Yaskawa INFORM job: 1C.JBI

/JOB
//NAME 1C
//POS
///NPOS 158,158,158,0,0,0
///TOOL 0
///POSTYPE PULSE
///PULSE
C00000=-283,-101162,-84213,3710,-80188,-1936
C00001=-283,-101162,-84213,3710,-80188,-1936
C00002=115939,-17843,-44700,-6904,-63515,59085
C00003=117851,11933,-44505,-6369,-54198,83131
C00004=117851,11880,-44474,-6366,-54245,83128
C00005=122172,13834,-42483,-463,-55485,73026
C00006=123748,7907,-48931,-483,-47630,63398
C00007=132704,14873,-45616,19438,-48261,40889
C00008=144175,42753,-30632,47438,-65070,14364
C00009=138306,51388,-15179,31478,-70676,13726
C00010=124819,56222,-2350,7571,-72880,2284
C00011=116170,53958,-4566,-7680,-71260,-3372
C00012=115645,53451,-5308,-7587,-71110,-3203
C00013=105039,58487,-7775,-25060,-77645,-21422
C00014=105262,24233,-38773,-26336,-58236,-42750
C00015=112386,11538,-46723,-12183,-49538,-53931
C00016=113021,10637,-47169,-12111,-49646,-54178
C00017=114170,-2374,-36949,-11645,-74681,-76938
C00018=113314,-7643,-38017,-11019,-76954,88145
C00019=103750,23668,-33240,-5111,-62302,87132
C00020=103750,23668,-33240,-5111,-62302,87132
C00021=110000,19960,-36933,2978,-58383,70645
C00022=112282,4054,-54561,4290,-38284,55376
C00023=127051,24932,-43086,41803,-51861,24110
C00024=126194,29403,-37517,40726,-52338,12802
C00025=118348,60362,-873,17694,-75878,15915
C00026=113933,56425,-1953,14226,-71232,-2232
C00027=100489,57495,-1416,-9321,-72833,-11727
C00028=101235,67629,7170,-3443,-84055,-29367
C00029=91022,64610,-2293,-23930,-82984,-31980
C00030=91048,41774,-22566,-24453,-68601,-40164
C00031=95890,27642,-32117,-16170,-61880,-54638
C00032=99594,19595,-38153,-13704,-58617,-69999
C00033=99594,19595,-38153,-13704,-58617,-69999
C00034=99303,8604,-31154,-10952,-72489,-71699
C00035=89422,16015,-23794,-2157,-75183,91094
C00036=91258,36004,-20905,-2546,-66652,90674
C00037=91258,36004,-20905,-2546,-66652,90674
C00038=96503,26815,-30375,3612,-58434,75085
C00039=104020,23579,-36756,17418,-51330,55937
C00040=113925,24192,-46060,50390,-45511,24597
C00041=112444,33459,-33623,40844,-50589,18382
C00042=105959,57894,-2087,19635,-69139,16595
C00043=102683,60172,2471,16804,-69167,938
C00044=91677,70980,13878,-1332,-78340,-10515
C00045=88699,81890,23139,-3974,-89133,-24557
C00046=80671,78616,14523,-19772,-88214,-29795
C00047=78063,59896,-4715,-24982,-77170,-36166
C00048=85285,24138,-35146,-12407,-50182,-52228
C00049=86525,30815,-27295,-12530,-61226,-65994
C00050=86525,30815,-27295,-12530,-61226,-65994
C00051=85063,22114,-18753,-9149,-74798,-67250
C00052=72786,31521,-9549,-9445,-75352,93043
C00053=79270,46324,-10095,-3085,-64870,94947
C00054=79270,46324,-10095,-3085,-64870,94947
C00055=83456,34403,-23445,1140,-53460,77595
C00056=88522,20590,-42092,13133,-33660,59513
C00057=92436,17350,-49768,33792,-25093,42436
C00058=100206,32488,-37788,50464,-41880,29044
C00059=99515,40284,-26338,41283,-46537,21581
C00060=98850,50643,-13462,39809,-52949,6831
C00061=91416,72483,16804,17125,-70588,4779
C00062=77894,87800,33476,-9278,-82729,-4550
C00063=79100,99899,45363,-1333,-94418,-21524
C00064=71782,98288,39798,-16226,-95116,-28048
C00065=67514,73380,11419,-25280,-78247,-32294
C00066=71390,53275,-6196,-18119,-65968,-46219
C00067=75669,46789,-10605,-11160,-64696,-62839
C00068=75669,46789,-10605,-11160,-64696,-62839
C00069=75039,37514,-3449,-7701,-77257,-64173
C00070=74616,28156,-12897,-9694,-74827,92488
C00071=75373,46749,-10374,-11505,-65177,93523
C00072=75373,46749,-10374,-11505,-65177,93523
C00073=83279,33454,-24235,1133,-53460,80094
C00074=88369,19506,-42835,13038,-33732,59606
C00075=92444,17438,-49755,33860,-25059,42415
C00076=100151,32274,-37986,50479,-41858,29056
C00077=99355,40003,-26600,41299,-46462,21619
C00078=100227,49460,-16867,46071,-52279,4034
C00079=91121,71677,16006,17029,-70030,4838
C00080=77993,87883,33867,-9296,-82912,-4592
C00081=79224,100354,46205,-1382,-94698,-21563
C00082=71921,98119,39548,-16283,-95028,-28080
C00083=67714,73606,11420,-25325,-78089,-32328
C00084=72711,51649,-6846,-14661,-65755,-51476
C00085=77715,33845,-23990,-6443,-52382,-64694
C00086=77715,33845,-23990,-6443,-52382,-64694
C00087=74844,35432,-1015,-7610,-79822,-64270
C00088=74616,28156,-12897,-9694,-74827,92488
C00089=90411,-2677,-20047,-11125,-84138,86440
C00090=90413,-2674,-20051,-11105,-84138,86441
C00091=137757,-12075,-30464,2646,-72394,74401
C00092=139263,-65150,-85436,14259,-28990,73053
C00093=136879,-25717,-69324,36252,-11746,62908
C00094=136879,-25717,-69324,36252,-11746,62908
C00095=139574,-23073,-65509,38333,-15951,40316
C00096=138446,-25572,-68856,45528,-10204,18708
C00097=136949,-21437,-61441,19475,-16251,9146
C00098=134482,-8675,-45493,4060,-31940,-3283
C00099=132921,-12133,-49426,2962,-29419,-26290
C00100=133351,-16693,-54684,5355,-25692,-47355
C00101=132569,-23850,-65218,-2678,-15038,-66834
C00102=133899,-27903,-74314,23479,-2636,-94546
C00103=138833,-79965,-103111,19688,-12213,-93629
C00104=119564,-93872,-103655,-3232,-19191,84847
C00105=119666,-28019,-68299,-3732,-15098,84700
C00106=119666,-28019,-68299,-3732,-15098,84700
C00107=119708,-30271,-73117,-29732,-7839,72372
C00108=119233,-27571,-67333,-20804,-14307,49665
C00109=119106,-25376,-64226,-16009,-16214,28430
C00110=118105,-24715,-63438,-17688,-16543,10280
C00111=116689,-17579,-54819,-12080,-26707,-16606
C00112=116486,-19327,-56780,-12438,-26446,-36213
C00113=109454,-19020,-60974,-47604,-29828,-43194
C00114=115085,-30409,-76062,-74083,-10783,-47674
C00115=113126,-78683,-102705,-45607,-16425,-60367
C00116=119564,-93872,-103655,-3232,-19191,84847
C00117=119355,-30239,-72733,-7438,-8938,86814
C00118=119355,-30239,-72733,-7438,-8938,86814
C00119=119373,-30935,-74214,-37542,-7197,75708
C00120=121407,-28868,-69424,-4086,-11316,43719
C00121=119107,-25533,-64139,-15884,-16345,28370
C00122=118122,-13860,-50139,-9217,-30457,5536
C00123=118283,-13038,-49068,-5042,-31449,-8478
C00124=116296,-14534,-51102,-10537,-31045,-19296
C00125=117896,-18615,-55611,-5957,-27309,-36360
C00126=112553,-24349,-66436,-46189,-21183,-44280
C00127=114320,-29666,-74035,-62528,-13006,-51221
C00128=113074,-79856,-103225,-44998,-16651,-60643
C00129=119564,-93872,-105617,-3232,-19191,84847
C00130=119652,-29586,-71182,-5048,-11389,85666
C00131=119652,-29586,-71182,-5048,-11389,85666
C00132=117863,-29049,-70076,-32838,-13629,71500
C00133=121453,-23804,-62042,-1822,-20367,42740
C00134=119106,-25569,-64361,-15996,-16232,28425
C00135=118129,-24991,-63785,-17715,-16469,10291
C00136=118320,-20483,-57910,-7080,-22477,-7740
C00137=116396,-17655,-54995,-12401,-26680,-16405
C00138=113643,-17458,-55850,-24185,-28054,-26576
C00139=114643,-26320,-67564,-36249,-17704,-47139
C00140=114895,-30423,-76085,-74235,-10895,-47569
C00141=112648,-89264,-107216,-40476,-18619,-62704
C00142=119564,-93872,-105617,-3232,-19191,84847
C00143=119574,-31211,-75378,-12278,-5097,88914
C00144=119574,-31211,-75378,-12278,-5097,88914
C00145=120258,-31594,-74917,-22580,-5990,69887
C00146=126376,-14543,-51553,17453,-33391,37954
C00147=119106,-25691,-64444,-15988,-16241,28420
C00148=117942,-25032,-63775,-18032,-16532,10469
C00149=116211,-17806,-55189,-12603,-26665,-16270
C00150=116661,-19498,-57018,-11750,-26290,-36065
C00151=116421,-21626,-59278,-15282,-26219,-55873
C00152=115105,-30520,-76064,-73793,-10790,-47808
C00153=112538,-91654,-108181,-39431,-19159,-63177
C00154=112538,-91654,-78834,-11871,-48570,95336
C00155=112538,-91654,-78834,-11871,-48570,95336
C00156=-2476,-84373,-75976,-13540,-83606,15477
C00157=-283,-101162,-84213,3710,-80188,-1936
BC00000=570125
BC00001=868704
BC00002=878894
BC00003=878037
BC00004=878037
BC00005=878038
BC00006=878038
BC00007=878038
BC00008=878038
BC00009=878038
BC00010=878038
BC00011=878038
BC00012=878038
BC00013=878038
BC00014=878037
BC00015=878037
BC00016=878037
BC00017=878037
BC00018=912823
BC00019=878035
BC00020=878035
BC00021=878037
BC00022=878037
BC00023=878038
BC00024=878037
BC00025=878038
BC00026=878038
BC00027=878037
BC00028=878037
BC00029=878037
BC00030=878037
BC00031=878037
BC00032=878037
BC00033=878037
BC00034=878037
BC00035=878035
BC00036=878036
BC00037=878036
BC00038=878037
BC00039=878037
BC00040=878038
BC00041=878038
BC00042=878038
BC00043=878038
BC00044=878037
BC00045=878037
BC00046=878037
BC00047=878037
BC00048=878037
BC00049=878037
BC00050=878037
BC00051=878037
BC00052=878037
BC00053=878035
BC00054=878035
BC00055=877203
BC00056=877947
BC00057=878201
BC00058=878342
BC00059=878784
BC00060=877961
BC00061=877604
BC00062=878505
BC00063=878840
BC00064=878535
BC00065=877953
BC00066=879795
BC00067=878428
BC00068=878428
BC00069=878037
BC00070=915550
BC00071=913919
BC00072=913919
BC00073=916409
BC00074=916569
BC00075=916479
BC00076=916387
BC00077=916586
BC00078=915550
BC00079=915870
BC00080=916359
BC00081=916889
BC00082=917058
BC00083=916344
BC00084=916666
BC00085=915811
BC00086=915811
BC00087=915811
BC00088=915550
BC00089=915550
BC00090=915550
BC00091=915550
BC00092=915550
BC00093=915550
BC00094=915550
BC00095=915550
BC00096=915550
BC00097=915550
BC00098=915550
BC00099=915550
BC00100=915550
BC00101=915550
BC00102=915550
BC00103=915550
BC00104=915550
BC00105=915551
BC00106=915551
BC00107=915550
BC00108=915550
BC00109=915550
BC00110=915550
BC00111=915550
BC00112=915550
BC00113=915550
BC00114=915550
BC00115=915550
BC00116=954211
BC00117=953187
BC00118=953187
BC00119=954162
BC00120=953948
BC00121=954071
BC00122=953633
BC00123=953445
BC00124=953244
BC00125=953645
BC00126=954029
BC00127=953749
BC00128=953683
BC00129=992214
BC00130=992214
BC00131=992214
BC00132=991968
BC00133=992423
BC00134=992186
BC00135=992082
BC00136=991590
BC00137=991168
BC00138=991569
BC00139=992735
BC00140=991845
BC00141=991844
BC00142=1026906
BC00143=1030289
BC00144=1030289
BC00145=1030261
BC00146=1030281
BC00147=1030485
BC00148=1029902
BC00149=1029299
BC00150=1030152
BC00151=1030177
BC00152=1030552
BC00153=1030552
BC00154=1030552
BC00155=1030552
BC00156=952617
BC00157=570125
EC00000=1164,0
EC00001=1166,0
EC00002=-1742,0
EC00003=-1741,0
EC00004=-1741,0
EC00005=-1742,0
EC00006=-1742,0
EC00007=-1741,0
EC00008=-1741,0
EC00009=-1741,0
EC00010=-1741,0
EC00011=-1741,0
EC00012=-1741,0
EC00013=-1742,0
EC00014=-1742,0
EC00015=-1742,0
EC00016=-1742,0
EC00017=-1741,0
EC00018=-1741,0
EC00019=-1744,0
EC00020=-1744,0
EC00021=-1742,0
EC00022=-1742,0
EC00023=-1741,0
EC00024=-1741,0
EC00025=-1741,0
EC00026=-1741,0
EC00027=-1741,0
EC00028=-1741,0
EC00029=-1742,0
EC00030=-1742,0
EC00031=-1741,0
EC00032=-1741,0
EC00033=-1741,0
EC00034=-1741,0
EC00035=-1743,0
EC00036=-1742,0
EC00037=-1742,0
EC00038=-1742,0
EC00039=-1742,0
EC00040=-1741,0
EC00041=-1741,0
EC00042=-1595,0
EC00043=-1742,0
EC00044=-1741,0
EC00045=-1741,0
EC00046=-1742,0
EC00047=-1742,0
EC00048=-1741,0
EC00049=-1741,0
EC00050=-1741,0
EC00051=-1741,0
EC00052=-1741,0
EC00053=-1743,0
EC00054=-1743,0
EC00055=-1742,0
EC00056=-1743,0
EC00057=-1742,0
EC00058=-1741,0
EC00059=-1741,0
EC00060=-1742,0
EC00061=-1742,0
EC00062=-1742,0
EC00063=-1741,0
EC00064=-1741,0
EC00065=-1741,0
EC00066=-1741,0
EC00067=-1742,0
EC00068=-1742,0
EC00069=-1741,0
EC00070=-1741,0
EC00071=-1742,0
EC00072=-1742,0
EC00073=-1742,0
EC00074=-1743,0
EC00075=-1742,0
EC00076=-1741,0
EC00077=-1740,0
EC00078=-1742,0
EC00079=-1742,0
EC00080=-1742,0
EC00081=-1741,0
EC00082=-1741,0
EC00083=-1741,0
EC00084=-1742,0
EC00085=-1742,0
EC00086=-1742,0
EC00087=-1741,0
EC00088=-1741,0
EC00089=-1741,0
EC00090=-84878,0
EC00091=-84879,0
EC00092=-84877,0
EC00093=-84877,0
EC00094=-84877,0
EC00095=-84877,0
EC00096=-84877,0
EC00097=-84877,0
EC00098=-84877,0
EC00099=-84877,0
EC00100=-84877,0
EC00101=-84877,0
EC00102=-84877,0
EC00103=-84877,0
EC00104=-84877,0
EC00105=-84878,0
EC00106=-84878,0
EC00107=-84877,0
EC00108=-84877,0
EC00109=-84877,0
EC00110=-84877,0
EC00111=-84877,0
EC00112=-84877,0
EC00113=-84877,0
EC00114=-84877,0
EC00115=-84877,0
EC00116=-84877,0
EC00117=-84878,0
EC00118=-84878,0
EC00119=-84877,0
EC00120=-84877,0
EC00121=-84877,0
EC00122=-84877,0
EC00123=-84877,0
EC00124=-84877,0
EC00125=-84877,0
EC00126=-84877,0
EC00127=-84877,0
EC00128=-84877,0
EC00129=-84877,0
EC00130=-84877,0
EC00131=-84877,0
EC00132=-84877,0
EC00133=-84877,0
EC00134=-84877,0
EC00135=-84877,0
EC00136=-84877,0
EC00137=-84877,0
EC00138=-84877,0
EC00139=-84877,0
EC00140=-84877,0
EC00141=-84877,0
EC00142=-84877,0
EC00143=-84877,0
EC00144=-84877,0
EC00145=-84877,0
EC00146=-84877,0
EC00147=-84877,0
EC00148=-84877,0
EC00149=-84877,0
EC00150=-84877,0
EC00151=-84877,0
EC00152=-84877,0
EC00153=-84877,0
EC00154=-84877,0
EC00155=-2299,0
EC00156=-193,0
EC00157=1164,0
//INST
///DATE 2025/01/31 19:46
///COMM OZZ
///ATTR SC,RW
///GROUP1 RB1,BS1
///GROUP2 ST1
NOP
MOVJ C00000 BC00000 VJ=70.00 DEC=20  +MOVJ EC00000 VJ=70.00
MOVJ C00001 BC00001 VJ=40.00 DEC=20  +MOVJ EC00001 VJ=40.00
MOVJ C00002 BC00002 VJ=70.00 DEC=20  +MOVJ EC00002 VJ=70.00
MOVJ C00003 BC00003 VJ=40.00 DEC=20  +MOVJ EC00003 VJ=70.00
MACRO1 MJ#(0) ARGF5
ARCON
MOVC C00004 BC00004 V=4.2 DEC=20  +MOVJ EC00004 VJ=70.00
MOVC C00005 BC00005 V=4.2 DEC=20  +MOVJ EC00005 VJ=30.00
MOVC C00006 BC00006 V=4.2 DEC=20  +MOVJ EC00006 VJ=30.00
MOVC C00007 BC00007 V=4.2 DEC=20  +MOVJ EC00007 VJ=30.00
MOVC C00008 BC00008 V=4.2 DEC=20  +MOVJ EC00008 VJ=30.00
MOVC C00009 BC00009 V=4.2 DEC=20  +MOVJ EC00009 VJ=30.00
MOVC C00010 BC00010 V=4.2 DEC=20  +MOVJ EC00010 VJ=30.00
MOVC C00011 BC00011 V=4.2 DEC=20  +MOVJ EC00011 VJ=30.00
MOVJ C00012 BC00012 VJ=25.00 DEC=20  +MOVJ EC00012 VJ=25.00
MOVC C00013 BC00013 V=4.2 DEC=20  +MOVJ EC00013 VJ=30.00
MOVC C00014 BC00014 V=4.2 DEC=20  +MOVJ EC00014 VJ=30.00
MOVC C00015 BC00015 V=4.2 DEC=20  +MOVJ EC00015 VJ=30.00
MOVC C00016 BC00016 V=4.2 DEC=20  +MOVJ EC00016 VJ=30.00
ARCOF
MOVJ C00017 BC00017 VJ=40.00 DEC=20  +MOVJ EC00017 VJ=40.00
MOVJ C00018 BC00018 VJ=70.00 DEC=20  +MOVJ EC00018 VJ=0.78
MOVJ C00019 BC00019 VJ=30.00 DEC=20  +MOVJ EC00019 VJ=0.78
ARCON
MOVC C00020 BC00020 V=4.2 DEC=20  +MOVJ EC00020 VJ=0.78
MOVC C00021 BC00021 V=4.2 DEC=20  +MOVJ EC00021 VJ=0.78
MOVC C00022 BC00022 V=4.2 DEC=20  +MOVJ EC00022 VJ=30.00
MOVC C00023 BC00023 V=4.2 DEC=20  +MOVJ EC00023 VJ=30.00
MOVC C00024 BC00024 V=5.8 DEC=20  +MOVJ EC00024 VJ=30.00
MOVC C00025 BC00025 V=4.2 DEC=20  +MOVJ EC00025 VJ=30.00
MOVC C00026 BC00026 V=4.2 DEC=20  +MOVJ EC00026 VJ=30.00
MOVC C00027 BC00027 V=4.2 DEC=20  +MOVJ EC00027 VJ=30.00
MOVC C00028 BC00028 V=4.2 DEC=20  +MOVJ EC00028 VJ=30.00
MOVC C00029 BC00029 V=4.2 DEC=20  +MOVJ EC00029 VJ=30.00
MOVC C00030 BC00030 V=4.2 DEC=20  +MOVJ EC00030 VJ=30.00
MOVC C00031 BC00031 V=4.2 DEC=20  +MOVJ EC00031 VJ=30.00
MOVC C00032 BC00032 V=4.2 DEC=20  +MOVJ EC00032 VJ=30.00
MOVJ C00033 BC00033 VJ=25.00 DEC=20  +MOVJ EC00033 VJ=30.00
ARCOF
MOVJ C00034 BC00034 VJ=30.00 DEC=20  +MOVJ EC00034 VJ=30.00
MOVJ C00035 BC00035 VJ=30.00 DEC=20  +MOVJ EC00035 VJ=30.00
MOVJ C00036 BC00036 VJ=30.00 DEC=20  +MOVJ EC00036 VJ=30.00
ARCON
MOVC C00037 BC00037 V=4.2 DEC=20  +MOVJ EC00037 VJ=30.00
MOVC C00038 BC00038 V=4.2 DEC=20  +MOVJ EC00038 VJ=30.00
MOVC C00039 BC00039 V=4.2 DEC=20  +MOVJ EC00039 VJ=30.00
MOVC C00040 BC00040 V=4.2 DEC=20  +MOVJ EC00040 VJ=30.00
MOVC C00041 BC00041 V=4.2 DEC=20  +MOVJ EC00041 VJ=30.00
MOVC C00042 BC00042 V=4.2 DEC=20  +MOVJ EC00042 VJ=30.00
MOVC C00043 BC00043 V=4.2 DEC=20  +MOVJ EC00043 VJ=30.00
MOVC C00044 BC00044 V=4.2 DEC=20  +MOVJ EC00044 VJ=30.00
MOVC C00045 BC00045 V=4.2 DEC=20  +MOVJ EC00045 VJ=30.00
MOVC C00046 BC00046 V=4.2 DEC=20  +MOVJ EC00046 VJ=30.00
MOVC C00047 BC00047 V=5.8 DEC=20  +MOVJ EC00047 VJ=30.00
MOVC C00048 BC00048 V=4.2 DEC=20  +MOVJ EC00048 VJ=0.78
MOVC C00049 BC00049 V=4.2 DEC=20  +MOVJ EC00049 VJ=30.00
MOVJ C00050 BC00050 VJ=30.00 DEC=20  +MOVJ EC00050 VJ=30.00
ARCOF
MOVJ C00051 BC00051 VJ=30.00 DEC=20  +MOVJ EC00051 VJ=30.00
MOVJ C00052 BC00052 VJ=30.00 DEC=20  +MOVJ EC00052 VJ=30.00
MOVJ C00053 BC00053 VJ=30.00 DEC=20  +MOVJ EC00053 VJ=30.00
ARCON
MOVC C00054 BC00054 V=4.2 DEC=20  +MOVJ EC00054 VJ=30.00
MOVC C00055 BC00055 V=4.2 DEC=20  +MOVJ EC00055 VJ=0.78
MOVC C00056 BC00056 V=4.2 DEC=20  +MOVJ EC00056 VJ=0.78
MOVC C00057 BC00057 V=4.2 DEC=20  +MOVJ EC00057 VJ=0.78
MOVC C00058 BC00058 V=4.2 DEC=20  +MOVJ EC00058 VJ=0.78
MOVC C00059 BC00059 V=4.2 DEC=20  +MOVJ EC00059 VJ=0.78
MOVC C00060 BC00060 V=4.2 DEC=20  +MOVJ EC00060 VJ=0.78
MOVC C00061 BC00061 V=4.2 DEC=20  +MOVJ EC00061 VJ=0.78
MOVC C00062 BC00062 V=4.2 DEC=20  +MOVJ EC00062 VJ=0.78
MOVC C00063 BC00063 V=4.2 DEC=20  +MOVJ EC00063 VJ=0.78
MOVC C00064 BC00064 V=4.2 DEC=20  +MOVJ EC00064 VJ=0.78
MOVC C00065 BC00065 V=4.2 DEC=20  +MOVJ EC00065 VJ=0.78
MOVC C00066 BC00066 V=4.2 DEC=20  +MOVJ EC00066 VJ=0.78
MOVC C00067 BC00067 V=4.2 DEC=20  +MOVJ EC00067 VJ=0.78
MOVJ C00068 BC00068 VJ=30.00 DEC=20  +MOVJ EC00068 VJ=30.00
ARCOF
MOVJ C00069 BC00069 VJ=30.00 DEC=20  +MOVJ EC00069 VJ=30.00
MOVJ C00070 BC00070 VJ=30.00 DEC=20  +MOVJ EC00070 VJ=30.00
MOVJ C00071 BC00071 VJ=30.00 DEC=20  +MOVJ EC00071 VJ=30.00
ARCON
MOVC C00072 BC00072 V=4.2 DEC=20  +MOVJ EC00072 VJ=30.00
MOVC C00073 BC00073 V=4.2 DEC=20  +MOVJ EC00073 VJ=30.00
MOVC C00074 BC00074 V=4.2 DEC=20  +MOVJ EC00074 VJ=30.00
MOVC C00075 BC00075 V=4.2 DEC=20  +MOVJ EC00075 VJ=40.00
MOVC C00076 BC00076 V=4.2 DEC=20  +MOVJ EC00076 VJ=30.00
MOVC C00077 BC00077 V=4.2 DEC=20  +MOVJ EC00077 VJ=25.00
MOVC C00078 BC00078 V=4.2 DEC=20  +MOVJ EC00078 VJ=30.00
MOVC C00079 BC00079 V=4.2 DEC=20  +MOVJ EC00079 VJ=70.00
MOVC C00080 BC00080 V=4.2 DEC=20  +MOVJ EC00080 VJ=30.00
MOVC C00081 BC00081 V=4.2 DEC=20  +MOVJ EC00081 VJ=30.00
MOVC C00082 BC00082 V=4.2 DEC=20  +MOVJ EC00082 VJ=30.00
MOVC C00083 BC00083 V=4.2 DEC=20  +MOVJ EC00083 VJ=30.00
MOVC C00084 BC00084 V=4.2 DEC=20  +MOVJ EC00084 VJ=0.78
MOVC C00085 BC00085 V=4.2 DEC=20  +MOVJ EC00085 VJ=30.00
MOVJ C00086 BC00086 VJ=25.00 DEC=20  +MOVJ EC00086 VJ=30.00
ARCOF
MOVJ C00087 BC00087 VJ=30.00 DEC=20  +MOVJ EC00087 VJ=30.00
MOVJ C00088 BC00088 VJ=30.00 DEC=20  +MOVJ EC00088 VJ=30.00
MOVJ C00089 BC00089 VJ=30.00 DEC=20  +MOVJ EC00089 VJ=30.00
MOVJ C00090 BC00090 VJ=30.00 DEC=20  +MOVJ EC00090 VJ=30.00
MOVJ C00091 BC00091 VJ=30.00 DEC=20  +MOVJ EC00091 VJ=30.00
MOVJ C00092 BC00092 VJ=70.00 DEC=20  +MOVJ EC00092 VJ=0.78
MOVJ C00093 BC00093 VJ=30.00 DEC=20  +MOVJ EC00093 VJ=0.78
MACRO1 MJ#(0) ARGF4
ARCON
MOVC C00094 BC00094 V=5.0 DEC=20  +MOVJ EC00094 VJ=0.78
MOVC C00095 BC00095 V=5.0 DEC=20  +MOVJ EC00095 VJ=0.78
MOVC C00096 BC00096 V=5.0 DEC=20  +MOVJ EC00096 VJ=0.78
MOVC C00097 BC00097 V=5.0 DEC=20  +MOVJ EC00097 VJ=0.78
MOVC C00098 BC00098 V=5.0 DEC=20  +MOVJ EC00098 VJ=0.78
MOVC C00099 BC00099 V=5.0 DEC=20  +MOVJ EC00099 VJ=0.78
MOVC C00100 BC00100 V=5.0 DEC=20  +MOVJ EC00100 VJ=0.78
MOVC C00101 BC00101 V=5.0 DEC=20  +MOVJ EC00101 VJ=0.78
MOVC C00102 BC00102 V=5.0 DEC=20  +MOVJ EC00102 VJ=0.78
ARCOF
MOVJ C00103 BC00103 VJ=40.00 DEC=20  +MOVJ EC00103 VJ=0.78
MOVJ C00104 BC00104 VJ=40.00 DEC=20  +MOVJ EC00104 VJ=0.78
MOVJ C00105 BC00105 VJ=40.00 DEC=20  +MOVJ EC00105 VJ=0.78
ARCON
MOVC C00106 BC00106 V=5.0 DEC=20  +MOVJ EC00106 VJ=0.78
MOVC C00107 BC00107 V=5.0 DEC=20  +MOVJ EC00107 VJ=0.78
MOVC C00108 BC00108 V=5.0 DEC=20  +MOVJ EC00108 VJ=40.00
MOVC C00109 BC00109 V=5.0 DEC=20  +MOVJ EC00109 VJ=0.78
MOVC C00110 BC00110 V=5.0 DEC=20  +MOVJ EC00110 VJ=0.78
MOVC C00111 BC00111 V=5.0 DEC=20  +MOVJ EC00111 VJ=0.78
MOVC C00112 BC00112 V=5.0 DEC=20  +MOVJ EC00112 VJ=0.78
MOVC C00113 BC00113 V=5.0 DEC=20  +MOVJ EC00113 VJ=0.78
MOVC C00114 BC00114 V=5.0 DEC=20  +MOVJ EC00114 VJ=0.78
ARCOF
MOVJ C00115 BC00115 VJ=40.00 DEC=20  +MOVJ EC00115 VJ=0.78
MOVJ C00116 BC00116 VJ=40.00 DEC=20  +MOVJ EC00116 VJ=0.78
MOVJ C00117 BC00117 VJ=40.00 DEC=20  +MOVJ EC00117 VJ=0.78
ARCON
MOVC C00118 BC00118 V=5.0 DEC=20  +MOVJ EC00118 VJ=0.78
MOVC C00119 BC00119 V=5.0 DEC=20  +MOVJ EC00119 VJ=0.78
MOVC C00120 BC00120 V=5.0 DEC=20  +MOVJ EC00120 VJ=0.78
MOVC C00121 BC00121 V=5.0 DEC=20  +MOVJ EC00121 VJ=0.78
MOVC C00122 BC00122 V=5.0 DEC=20  +MOVJ EC00122 VJ=0.78
MOVC C00123 BC00123 V=5.0 DEC=20  +MOVJ EC00123 VJ=0.78
MOVC C00124 BC00124 V=5.0 DEC=20  +MOVJ EC00124 VJ=0.78
MOVC C00125 BC00125 V=5.0 DEC=20  +MOVJ EC00125 VJ=0.78
MOVC C00126 BC00126 V=5.0 DEC=20  +MOVJ EC00126 VJ=0.78
MOVC C00127 BC00127 V=5.0 DEC=20  +MOVJ EC00127 VJ=0.78
ARCOF
MOVJ C00128 BC00128 VJ=40.00 DEC=20  +MOVJ EC00128 VJ=0.78
MOVJ C00129 BC00129 VJ=40.00 DEC=20  +MOVJ EC00129 VJ=0.78
MOVJ C00130 BC00130 VJ=40.00 DEC=20  +MOVJ EC00130 VJ=0.78
ARCON
MOVC C00131 BC00131 V=5.0 DEC=20  +MOVJ EC00131 VJ=0.78
MOVC C00132 BC00132 V=5.0 DEC=20  +MOVJ EC00132 VJ=0.78
MOVC C00133 BC00133 V=5.0 DEC=20  +MOVJ EC00133 VJ=0.78
MOVC C00134 BC00134 V=5.0 DEC=20  +MOVJ EC00134 VJ=0.78
MOVC C00135 BC00135 V=5.0 DEC=20  +MOVJ EC00135 VJ=0.78
MOVC C00136 BC00136 V=5.0 DEC=20  +MOVJ EC00136 VJ=0.78
MOVC C00137 BC00137 V=5.0 DEC=20  +MOVJ EC00137 VJ=0.78
MOVC C00138 BC00138 V=5.0 DEC=20  +MOVJ EC00138 VJ=0.78
MOVC C00139 BC00139 V=5.0 DEC=20  +MOVJ EC00139 VJ=0.78
MOVC C00140 BC00140 V=5.0 DEC=20  +MOVJ EC00140 VJ=0.78
ARCOF
MOVJ C00141 BC00141 VJ=40.00 DEC=20  +MOVJ EC00141 VJ=0.78
MOVJ C00142 BC00142 VJ=40.00 DEC=20  +MOVJ EC00142 VJ=0.78
MOVJ C00143 BC00143 VJ=40.00 DEC=20  +MOVJ EC00143 VJ=0.78
ARCON
MOVC C00144 BC00144 V=5.0 DEC=20  +MOVJ EC00144 VJ=0.78
MOVC C00145 BC00145 V=5.0 DEC=20  +MOVJ EC00145 VJ=0.78
MOVC C00146 BC00146 V=5.0 DEC=20  +MOVJ EC00146 VJ=0.78
MOVC C00147 BC00147 V=5.0 DEC=20  +MOVJ EC00147 VJ=0.78
MOVC C00148 BC00148 V=5.0 DEC=20  +MOVJ EC00148 VJ=0.78
MOVC C00149 BC00149 V=5.0 DEC=20  +MOVJ EC00149 VJ=0.78
MOVC C00150 BC00150 V=5.0 DEC=20  +MOVJ EC00150 VJ=0.78
MOVC C00151 BC00151 V=5.0 DEC=20  +MOVJ EC00151 VJ=0.78
MOVC C00152 BC00152 V=5.0 DEC=20  +MOVJ EC00152 VJ=0.78
ARCOF
MOVJ C00153 BC00153 VJ=40.00 DEC=20  +MOVJ EC00153 VJ=0.78
MOVJ C00154 BC00154 VJ=40.00 DEC=20  +MOVJ EC00154 VJ=0.78
MOVJ C00155 BC00155 VJ=40.00 DEC=20  +MOVJ EC00155 VJ=40.00
MOVJ C00156 BC00156 VJ=40.00 DEC=20  +MOVJ EC00156 VJ=0.78
MOVJ C00157 BC00157 VJ=40.00 DEC=20  +MOVJ EC00157 VJ=0.78
END
